Fanuc KAREL source: kb00171.KL

-- PROVISIONAL review KL for V1013-1; original PC SHA256 0eb25450bb065b2070a6ce04a200b93bfcbbc4ba3753e9e2547df660f976c991
-- Incomplete behavior may be omitted. Consult companion uncertainty JSON. Do not deploy.
PROGRAM KB00171
%NOLOCKGROUP
BEGIN
  -- UNRESOLVED_PC offsets 5-12; opcodes 9D,23
  -- UNRESOLVED_PC offsets 17-24; opcodes 9D,23
  -- UNRESOLVED_PC offsets 29-36; opcodes 9D,23
  -- UNRESOLVED_PC offsets 41-69; opcodes 27,22,22,22,31,23
  -- UNRESOLVED_PC offsets 74-78; opcodes 7F
END KB00171
